(* IEC 61131-3 sources: IRIS-Project/LASAL CONTROL SOFTWARE/LasalProject_2025_09_12/Class/IrradiationManager, 1 file *)

(* ---- IrradiationManager.st ---- *)
(*!
<Class
	Name               = "IrradiationManager"
	Revision           = "0.0"
	RealtimeTask       = "false"
	CyclicTask         = "true"
	DefCyclictime      = "100 ms"
	BackgroundTask     = "false"
	Sigmatek           = "false"
	OSInterface        = "false"
	HighPriority       = "false"
	Automatic          = "false"
	UpdateMode         = "Prescan"
	SharedCommandTable = "true"
	Objectsize         = "(560,120)">
	<Channels>
		<Server Name="ClassSvr" Visualized="false" Initialize="false" WriteProtected="true" Retentive="false"/>
		<Server Name="s_1_3_pelletMode" Visualized="false" Initialize="false" WriteProtected="false" Retentive="false"/>
		<Server Name="s_EasyGUI" Visualized="false" Initialize="false" WriteProtected="false" Retentive="false"/>
		<Server Name="s_Reset" Visualized="false" Initialize="false" WriteProtected="false" Retentive="false"/>
		<Server Name="s_setTimer1" Visualized="false" Initialize="false" WriteProtected="false" Retentive="false"/>
		<Server Name="s_setTimer2" Visualized="false" Initialize="false" WriteProtected="false" Retentive="false"/>
		<Server Name="s_setTimer3" Visualized="false" Initialize="false" WriteProtected="false" Retentive="false"/>
		<Server Name="s_TimerStartStop" Visualized="false" Initialize="false" WriteProtected="false" Retentive="false"/>
		<Server Name="s_VisTimerIrr1" Visualized="false" Initialize="false" WriteProtected="false" Retentive="false"/>
		<Server Name="s_VisTimerIrr2" Visualized="false" Initialize="false" WriteProtected="false" Retentive="false"/>
		<Server Name="s_VisTimerIrr3" Visualized="false" Initialize="false" WriteProtected="false" Retentive="false"/>
		<Server Name="s_VisTimerIrrAdv1" Visualized="false" Initialize="false" WriteProtected="false" Retentive="false"/>
		<Server Name="s_VisTimerIrrAdv2" Visualized="false" Initialize="false" WriteProtected="false" Retentive="false"/>
		<Server Name="s_VisTimerIrrAdv3" Visualized="false" Initialize="false" WriteProtected="false" Retentive="false"/>
		<Server Name="Startprocess" Visualized="false" Initialize="false" WriteProtected="false" Retentive="false"/>
		<Client Name="c_SysTime" Required="true" Internal="false"/>
		<Client Name="c_timerLib" Required="true" Internal="false"/>
		<Client Name="NrIrrTablets" Required="true" Internal="false"/>
		<Client Name="SetStartStopIrr" Required="true" Internal="false"/>
		<Client Name="TabletInIrrPos" Required="true" Internal="false"/>
		<Client Name="Timer1" Required="true" Internal="false"/>
		<Client Name="Timer2" Required="true" Internal="false"/>
		<Client Name="Timer3" Required="true" Internal="false"/>
	</Channels>
	<Separators>
		<Servers>
			<SepChn Position="8"/>
			<SepChn Position="4"/>
			<SepChn Position="12"/>
		</Servers>
		<Clients>
			<SepChn Position="3"/>
			<SepChn Position="6"/>
		</Clients>
	</Separators>
</Class>
*)
IrradiationManager : CLASS
	TYPE
	  t_timerCase :  //! <Type Public="true" Name="t_timerCase"/>
	  (
	    Idle:=30,
	    tablet1:=0,
	    tablet2:=10,
	    tablet3:=20
	  )$UDINT;
	END_TYPE
  //Servers:
	ClassSvr 	: SvrChCmd_DINT;
	s_setTimer1 	: SvrCh_UDINT;
	s_setTimer2 	: SvrCh_UDINT;
	s_setTimer3 	: SvrCh_UDINT;
	s_VisTimerIrr1 	: SvrCh_UDINT;
	s_VisTimerIrr2 	: SvrCh_UDINT;
	s_VisTimerIrr3 	: SvrCh_UDINT;
	s_VisTimerIrrAdv1 	: SvrCh_DINT;
	s_VisTimerIrrAdv2 	: SvrCh_DINT;
	s_VisTimerIrrAdv3 	: SvrCh_DINT;
	Startprocess 	: SvrCh_DINT;
	s_EasyGUI 	: SvrCh_DINT;
	s_Reset 	: SvrCh_DINT;
	s_TimerStartStop 	: SvrCh_DINT;
	s_1_3_pelletMode 	: SvrCh_DINT;
  //Clients:
	Timer1 	: CltChCmd_TimerLib;
	Timer2 	: CltChCmd_TimerLib;
	Timer3 	: CltChCmd_TimerLib;
	TabletInIrrPos 	: CltCh_DINT;
	NrIrrTablets 	: CltCh_DINT;
	SetStartStopIrr 	: CltCh_t_IrradiationPhase_PTofCls_Manager_globale;
	c_timerLib 	: CltChCmd_TimeDateLib;
	c_SysTime 	: CltCh_TIME_LSL;
  //Variables:
		v_StartProcess 	: DINT;
		v_NrTablets 	: DINT;
		v_TabletInIrrPos 	: DINT;
		v_Timer1 	: UDINT;
		v_Timer2 	: UDINT;
		v_Timer3 	: UDINT;
		c_CaseTimer 	: DINT;
		c_Timer1 	: DINT;
		c_Timer2 	: DINT;
		c_Timer3 	: DINT;
		startTimer1 	: UDINT;
		startTimer2 	: UDINT;
		startTimer3 	: UDINT;
		v_startCases 	: DINT;
		v_EasyGUI 	: DINT;
		v_hd_Time_1 	: HDINT;
		v_hd_Time_2 	: HDINT;
		v_tot_seconds 	: DINT;
  //Functions:

	FUNCTION VIRTUAL GLOBAL Init;

	FUNCTION VIRTUAL GLOBAL CyWork
		VAR_INPUT
			EAX 	: UDINT;
		END_VAR
		VAR_OUTPUT
			state (EAX) 	: UDINT;
		END_VAR;

	FUNCTION VIRTUAL GLOBAL Startprocess::Read
		VAR_OUTPUT
			output (EAX) 	: DINT;
		END_VAR;

	FUNCTION VIRTUAL GLOBAL s_EasyGUI::Read
		VAR_OUTPUT
			output (EAX) 	: DINT;
		END_VAR;
  //Tables:
	FUNCTION @STD
		VAR_OUTPUT
			ret_code	: CONFSTATES;
		END_VAR;
	FUNCTION GLOBAL TAB @CT_;
END_CLASS;

#pragma usingLtd TimeDateLib
#pragma usingLtd TimerLib

FUNCTION VIRTUAL GLOBAL IrradiationManager::CyWork
	VAR_INPUT
		EAX 	: UDINT;
	END_VAR
	VAR_OUTPUT
		state (EAX) 	: UDINT;
	END_VAR

//set Timer dai server
v_Timer1:=1000*s_setTimer1;
v_Timer2:=1000*s_setTimer2;
v_Timer3:=1000*s_setTimer3;

//get status of tablet (irr pos): Nr and position
v_TabletInIrrPos:=TabletInIrrPos.Read();
v_NrTablets:=NrIrrTablets.Read();

v_EasyGUI:=s_EasyGUI.Read();

v_StartProcess:=Startprocess.Read();

  if s_Reset.Read() then
     s_VisTimerIrr1.Write(input:=0);
     s_VisTimerIrr2.Write(input:=0);
     s_VisTimerIrr3.Write(input:=0);
     s_VisTimerIrrAdv1.Write(input:=0);
     s_VisTimerIrrAdv2.Write(input:=0);
     s_VisTimerIrrAdv3.Write(input:=0);
     c_Timer1:=0;
     c_Timer2:=0;
     c_Timer3:=0;
     c_CaseTimer:=30;
     startTimer1:=0;
     startTimer2:=0;
     startTimer3:=0;
     v_NrTablets:=0;
     s_setTimer1.Write(input:=0);
     s_setTimer2.Write(input:=0);
     s_setTimer3.Write(input:=0);
     Startprocess.Write(input:=0);

  end_if;

  if c_Timer3=30 & c_CaseTimer=20 then
    s_VisTimerIrr3.Write(input:=v_Timer3);
  end_if;

  if v_StartProcess & v_TabletInIrrPos & v_EasyGUI then

  case c_CaseTimer of

    30:
      c_CaseTimer:=10*v_NrTablets;
      v_startCases:=10;

    40:
      s_VisTimerIrr1.Write(input:=v_Timer1);

    0:

      case c_Timer1 of
        0:
          c_Timer1:=v_startCases;

        10:
          v_startCases:=0;
          Timer1.TimerStart(pudStartTime:=#startTimer1);
          SetStartStopIrr.Write(input:=Manager_globale::Irradiation_Start);
          c_Timer1:=20;

        20:
          if Timer1.IsTimerFinished(pudStartTime:=#startTimer1, udDuration:=v_Timer1) then
            SetStartStopIrr.Write(input:=Manager_globale::Irradiation_Over);
            c_CaseTimer:=30;
          end_if;

          s_VisTimerIrr1.Write(input:=Timer1.TimerRest(pudStartTime:=#startTimer1, udDuration:=v_Timer1));

      end_case;

    10:

       case c_Timer2 of
        0:
          c_Timer2:=v_startCases;
          s_VisTimerIrr1.Write(input:=v_Timer1);

        10:
          v_startCases:=0;
          Timer2.TimerStart(pudStartTime:=#startTimer2);
          SetStartStopIrr.Write(input:=Manager_globale::Irradiation_Start);
          c_Timer2:=20;

        20:
          if Timer2.IsTimerFinished(pudStartTime:=#startTimer2, udDuration:=v_Timer2) then
            SetStartStopIrr.Write(input:=Manager_globale::Irradiation_Over);
            c_CaseTimer:=30;
          end_if;

          s_VisTimerIrr2.Write(input:=Timer2.TimerRest(pudStartTime:=#startTimer2, udDuration:=v_Timer2));

      end_case;

    20:

      case c_Timer3 of
        0:
          c_Timer3:=v_startCases;
          s_VisTimerIrr2.Write(input:=v_Timer2);

        10:
          v_startCases:=0;
          Timer3.TimerStart(pudStartTime:=#startTimer3);
          SetStartStopIrr.Write(input:=Manager_globale::Irradiation_Start);
          c_Timer3:=20;

        20:
          if Timer3.IsTimerFinished(pudStartTime:=#startTimer3, udDuration:=v_Timer3) then
            SetStartStopIrr.Write(input:=Manager_globale::Irradiation_Over);
            c_Timer3:=30;
          end_if;

          s_VisTimerIrr3.Write(input:=Timer3.TimerRest(pudStartTime:=#startTimer3, udDuration:=v_Timer3));

         30:
          s_VisTimerIrr3.Write(input:=v_Timer3);

      end_case;

  end_case;

  elsif v_EasyGUI=0 then

    case c_CaseTimer of

    30:
      c_CaseTimer:=10*v_NrTablets;
      v_startCases:=10;

    0:

      case c_Timer1 of
        0:
          c_Timer1:=v_startCases;

        10:
          if s_TimerStartStop.Read() then
            v_hd_Time_1:=c_SysTime.Read();
            c_Timer1:=20;
          end_if;

        20:
          if s_TimerStartStop.Read()=0 then
            v_hd_Time_2:=c_SysTime.Read();
            c_Timer1:=30;
          end_if;

        30:
          v_tot_seconds := c_timerLib.TimeDiff(tim1:=v_hd_Time_2, tim2:=v_hd_Time_1);
          s_VisTimerIrrAdv1.Write(input:=v_tot_seconds);
          c_CaseTimer:=30;

      end_case;

    10:

       case c_Timer2 of
        0:
          c_Timer2:=v_startCases;

        10:
          if s_TimerStartStop.Read() then
            v_hd_Time_1:=c_SysTime.Read();
            c_Timer2:=20;
          end_if;

        20:
          if s_TimerStartStop.Read()=0 then
            v_hd_Time_2:=c_SysTime.Read();
            c_Timer2:=30;
          end_if;

        30:
          v_tot_seconds := c_timerLib.TimeDiff(tim1:=v_hd_Time_2, tim2:=v_hd_Time_1);
          s_VisTimerIrrAdv2.Write(input:=v_tot_seconds);
          c_CaseTimer:=30;

      end_case;

    20:

      case c_Timer3 of
        0:
          c_Timer3:=v_startCases;

        10:
          if s_TimerStartStop.Read() then
            v_hd_Time_1:=c_SysTime.Read();
            c_Timer3:=20;
          end_if;

        20:
          if s_TimerStartStop.Read()=0 then
            v_hd_Time_2:=c_SysTime.Read();
            c_Timer3:=30;
          end_if;

        30:
          v_tot_seconds := c_timerLib.TimeDiff(tim1:=v_hd_Time_2, tim2:=v_hd_Time_1);
          s_VisTimerIrrAdv3.Write(input:=v_tot_seconds);
          c_CaseTimer:=40;

        40:

      end_case;

    end_case;

  elsif v_EasyGUI=1 & s_1_3_pelletMode.Read()=1 & c_Timer1=20 then
     s_VisTimerIrr1.Write(input:=v_Timer1);

  end_if;

	state := READY;

END_FUNCTION

FUNCTION VIRTUAL GLOBAL IrradiationManager::Init

v_Timer1:=0;
v_Timer2:=0;
v_Timer3:=0;

v_TabletInIrrPos:=0;
v_NrTablets:=0;

v_StartProcess:=0;

c_Timer1:=0;
c_Timer2:=0;
c_Timer3:=0;

v_startCases:=0;

c_CaseTimer:=30;

v_EasyGUI:=0;

END_FUNCTION

FUNCTION VIRTUAL GLOBAL IrradiationManager::Startprocess::Read
	VAR_OUTPUT
		output (EAX) 	: DINT;
	END_VAR

	output := Startprocess;

END_FUNCTION

FUNCTION VIRTUAL GLOBAL IrradiationManager::s_EasyGUI::Read
	VAR_OUTPUT
		output (EAX) 	: DINT;
	END_VAR

	output := s_EasyGUI;

END_FUNCTION
